FUNCTION_BLOCK FB_RTC_1
VAR_INPUT
END_VAR
VAR_OUTPUT
	(* Variables *)
	bTimeValid							:BOOL;
	dtRTC        						:DT;
	dtRTCEX      						:DT;
	stDateTime							:ST_DateTime;
END_VAR
VAR
	(* Enummerations *)
	
	(* Variables *)
	bFirstTime							:BOOL;	
	bBusy								:BOOL;
	bError								:BOOL;
	udnErrorNo							:UDINT;			

	actSysTimeDate						:TIMESTRUCT;				(* Structure SysTimeDate *)
	
	bValidRTC      						:BOOL;	
	bValidRTCEX    						:BOOL;

	(* References *)

	(* Interfaces *)

	(* Instances *)

   	fbGetLocalTime  					:NT_GetTime;
	tonSyncTimer       					:TON;
	ftSyncTrigger     					:F_TRIG;

	rtFirstTime						:R_TRIG;

	fbRTC           						:RTC;
	fbRTCEX        						:RTC_EX;

	(* Information given by the RTC *)
	wYear								:WORD;
	wMonth								:WORD;
	wDay								:WORD;
	wHour								:WORD;
	wMinute								:WORD;
	wSecond							:WORD;
	wMilliseconds						:WORD;
	
	dtDatTimePunktHilfv :STRING;

END_VAR


IF NOT bFirstTime
THEN
	bFirstTime := TRUE;
	
END_IF


(* Get RTC *)
rtFirstTime(CLK := bFirstTime);

(* Time synchronization *)
tonSyncTimer(
	IN := NOT tonSyncTimer.Q,
	PT := T#100MS,
);

(* This function provides the time (seconds) which has passed since 01.01.1970 00:00:00 (RTC). *)
fbGetLocalTime(
	NETID := '',
	START := tonSyncTimer.Q
			 OR rtFirstTime.Q,
	TMOUT := T#5S,
	BUSY => bBusy,
	ERR => bError,
	ERRID => udnErrorNo
);

actSysTimeDate := fbGetLocalTime.TIMESTR;

(*This function converts the time given into format SysTimeDate.*)
ftSyncTrigger(CLK := bBusy AND NOT bError);

fbRTC(
	EN := ftSyncTrigger.Q, 
	PDT := SYSTEMTIME_TO_DT(actSysTimeDate), 
	Q => bValidRTC, 
	CDT => dtRTC 
);

fbRTCEX(
	EN := ftSyncTrigger.Q,
	PDT := SYSTEMTIME_TO_DT(actSysTimeDate),
	PMSEK := actSysTimeDate.wMilliseconds,
	Q => bValidRTCEX, 
	CDT => dtRTCEX 
);

(*The structure SysTimeDate contains detailed information on the system time, 
split up into a readable format, e.g.:*)

wYear := actSysTimeDate.wYear;
wMonth := actSysTimeDate.wMonth;
wDay := actSysTimeDate.wDay;
wHour := actSysTimeDate.wHour;
wMinute := actSysTimeDate.wMinute;
wSecond := actSysTimeDate.wSecond;
wMilliseconds := actSysTimeDate.wMilliseconds;

stDateTime.dtDateTime := dtRTC;
stDateTime.dtDateTimeEx := dtRTCEX;

stDateTime.sDate := CONCAT(WORD_TO_STRING(wYear),
		 CONCAT(SEL(LEN(WORD_TO_STRING(wMonth))=1 ,WORD_TO_STRING(wMonth),CONCAT('0',WORD_TO_STRING(wMonth))),
				SEL(LEN(WORD_TO_STRING(wDay))=1 ,WORD_TO_STRING(wDay),CONCAT('0',WORD_TO_STRING(wDay)))));

stDateTime.sTime := CONCAT(SEL(LEN(WORD_TO_STRING(wHour))=1 ,WORD_TO_STRING(wHour),CONCAT('0',WORD_TO_STRING(wHour))),
		 CONCAT(SEL(LEN(WORD_TO_STRING(wMinute))=1 ,WORD_TO_STRING(wMinute),CONCAT('0',WORD_TO_STRING(wMinute))),
				SEL(LEN(WORD_TO_STRING(wSecond))=1 ,WORD_TO_STRING(wSecond),CONCAT('0',WORD_TO_STRING(wSecond)))));

stDateTime.sTimeEx := CONCAT(stDateTime.sTime, SEL(LEN(WORD_TO_STRING(wMilliseconds))=1 , SEL(LEN(WORD_TO_STRING(wMilliseconds))=2 , WORD_TO_STRING(wMilliseconds), CONCAT('0',WORD_TO_STRING(wMilliseconds))), CONCAT('00',WORD_TO_STRING(wMilliseconds))));
				
stDateTime.sDateTime := CONCAT(stDateTime.sDate,CONCAT('_', stDateTime.sTime));

stDateTime.sDateTimeEx := CONCAT(stDateTime.sDate,CONCAT('_', stDateTime.sTimeEx));


dtDatTimePunktHilfv := DELETE(DT_TO_STRING(stDateTime.dtDateTime),4,0);
stDateTime.dtDateTimePunkt :=REPLACE(dtDatTimePunktHilfv,' ',1,11);

END_FUNCTION_BLOCK

(* stored: Version 1.1.0.1, ProductVersion 3.1.4024.15
   POU FB_RTC_1: Id {177c10ed-33c8-4fc6-ae89-7385ff72734d}, SpecialFunc None *)
